TYPE "ST_InnerUnitHal"
VERSION : 0.1
   STRUCT
      "Cell" {ExternalAccessible := 'False'; ExternalVisible := 'False'; ExternalWritable := 'False'} : "ST_DeclarationCellHal";
   END_STRUCT;
END_TYPE
